Fanuc KAREL source: KA00193.KL

PROGRAM KA00193
%NOLOCKGROUP
VAR
  SRC: ARRAY[4] OF SHORT
  DST: ARRAY[4] OF STRING[20]
BEGIN
  DST = SRC
END KA00193
